// This function has been automatically generated from the project information.
{attribute 'signature_flag' := '1073741824'}
{attribute 'TcGenerated'}
{attribute 'no-analysis'}
FUNCTION F_GetTitle : WSTRING
VAR_INPUT
	
END_VAR

F_GetTitle := "Intecre.TwinSAFE.Models";

END_FUNCTION

(* stored: Version 1.1.0.1
   POU F_GetTitle: Id {fa60f0ba-5d15-4aed-9391-fbc7f753d8bd}, SpecialFunc None *)
